Fanuc KAREL source: kt00579.KL

-- PROVISIONAL review KL for V940-1; original PC SHA256 a64810749bf3fffa5f2dbf9179633a8adc45f370e1be59aed6aac721f54cd7d1
-- Incomplete behavior may be omitted. Consult companion uncertainty JSON. Do not deploy.
PROGRAM KT00579
%NOLOCKGROUP
VAR
  I2 : INTEGER
-- UNRESOLVED_DECL V1 type=000013
-- UNRESOLVED_DECL OUT type=000013
BEGIN
  -- V9_ZERO_TABLE_METADATA_HINT layout=0001; no indexed target words; source/name/runtime held
  -- UNRESOLVED_PC offsets 5-20; opcodes 2E,22,32,35
  -- UNRESOLVED_PC offsets 25-36; opcodes 2E,23
  -- UNRESOLVED_PC offsets 41-63; opcodes 49,21,89,4A
  -- UNRESOLVED_PC offsets 68-72; opcodes 7F
END KT00579
